Yaskawa INFORM job: STAR.JBI

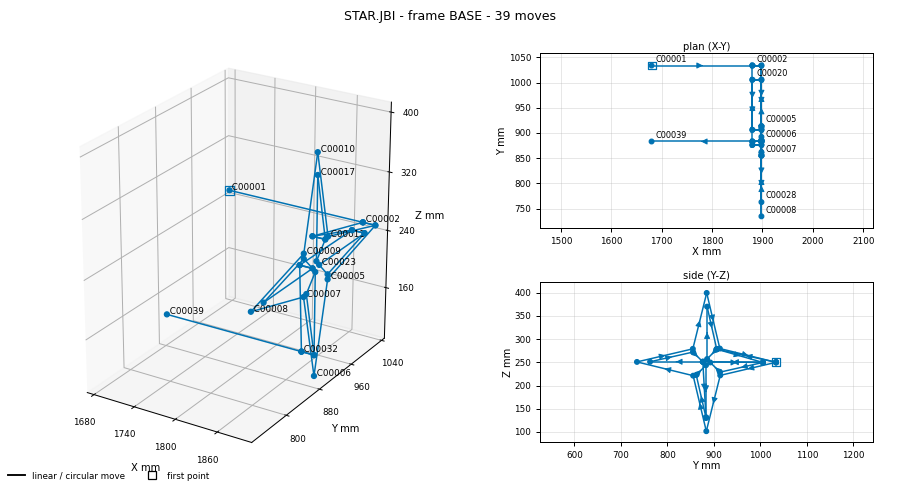
[picture p0: tool path of STAR.JBI in frame BASE, 39 of 40 moves have a stored position in this frame; points joined in program order, loops and branches not executed]
/JOB
//NAME STAR
//POS
///NPOS 40,0,0,0,0,0
///TOOL 9
///POSTYPE PULSE
///PULSE
C00000=38,23,-28,-44,61,-64
///TOOL 9
///POSTYPE BASE
///RECTAN
///RCONF 1,0,0,0,0,0,0,0
C00001=1680.000,1033.806,249.952,-90.00,-0.00,-90.00
C00002=1880.000,1033.806,249.952,-90.00,-0.00,-90.00
C00003=1880.000,1033.806,249.952,-90.00,-0.00,-90.00
C00004=1898.000,1033.806,249.952,-90.00,-0.00,-90.00
C00005=1898.000,913.725,221.863,-90.00,-0.00,-90.00
C00006=1898.000,883.747,101.722,-90.00,-0.00,-90.00
C00007=1898.000,855.472,221.186,-90.00,-0.00,-90.00
C00008=1898.000,734.538,250.798,-90.00,-0.00,-90.00
C00009=1898.000,854.791,278.888,-90.00,-0.00,-90.00
C00010=1898.000,884.598,399.198,-90.00,-0.00,-90.00
C00011=1898.000,912.873,279.564,-90.00,-0.00,-90.00
C00012=1898.000,1033.806,249.952,-90.00,-0.00,-90.00
C00013=1880.000,1033.806,249.952,-90.00,-0.00,-90.00
C00014=1880.000,906.230,278.211,-90.00,-0.00,-90.00
C00015=1898.000,906.230,278.211,-90.00,-0.00,-90.00
C00016=1898.000,885.450,257.059,-90.00,-0.00,-90.00
C00017=1898.000,885.450,369.755,-90.00,-0.00,-90.00
C00018=1898.000,906.230,278.211,-90.00,-0.00,-90.00
C00019=1880.000,906.230,278.211,-90.00,-0.00,-90.00
C00020=1880.000,1005.532,249.614,-90.00,-0.00,-90.00
C00021=1898.000,1005.532,249.614,-90.00,-0.00,-90.00
C00022=1898.000,913.384,228.801,-90.00,-0.00,-90.00
C00023=1898.000,892.263,249.614,-90.00,-0.00,-90.00
C00024=1898.000,1005.532,249.614,-90.00,-0.00,-90.00
C00025=1880.000,1005.532,249.614,-90.00,-0.00,-90.00
C00026=1880.000,876.252,251.137,-90.00,-0.00,-90.00
C00027=1898.000,876.252,251.137,-90.00,-0.00,-90.00
C00028=1898.000,762.813,251.137,-90.00,-0.00,-90.00
C00029=1898.000,854.961,271.950,-90.00,-0.00,-90.00
C00030=1898.000,876.252,251.137,-90.00,-0.00,-90.00
C00031=1880.000,876.252,251.137,-90.00,-0.00,-90.00
C00032=1880.000,883.065,130.996,-90.00,-0.00,-90.00
C00033=1898.000,883.065,130.996,-90.00,-0.00,-90.00
C00034=1898.000,862.115,222.540,-90.00,-0.00,-90.00
C00035=1898.000,883.065,243.691,-90.00,-0.00,-90.00
C00036=1898.000,883.065,130.996,-90.00,-0.00,-90.00
C00037=1880.000,883.065,130.996,-90.00,-0.00,-90.00
C00038=1880.000,883.065,130.996,-90.00,-0.00,-90.00
C00039=1680.000,883.065,130.996,-90.00,-0.00,-90.00
//INST
///DATE 2026/10/26 01:19
///COMM Generated using RoboDK
///ATTR SC,RW,RJ
///GROUP1 RB1
NOP
'Using Tool3 (targets wrt base
'):
'1900.0,883.5,250.0,90.0,0.0,-
'90.0
'Setting Tool 9 (USER - CONE -
' 10MM  X  45 DEG):
SETE P00095 (1) 0
SETE P00095 (2) 0
SETE P00095 (3) 85000
SETE P00095 (4) 0
SETE P00095 (5) 0
SETE P00095 (6) 0
SETTOOL TL#(9) P00095
'hide BALL END - 10MM
'show USER - CONE - 10MM  X  4
'5 DEG
MSG "/ ALPHACAM DRAWING FILE -"
MSG " ROBOTAPT"
MSG "/ NC CODE FILE - ROBOTAPT"
MSG ".apt"
MSG "/ POST-PROCESSED FOR APT-"
MSG "CL DATA"
MSG "/ CREATED - 26 NOV 18"
MSG "/ PROGRAMMED BY ALPHACAM"
MSG "/ USER - CONE - 10MM  X  "
MSG "45 DEG"
MOVJ C00000 VJ=50.00
MOVL C00001 V=1000.0
MOVL C00002 V=1000.0
CALL JOB:SPINDLE
MOVL C00003 V=1000.0
MOVL C00004 V=160.0
MOVL C00005 V=160.0
MOVL C00006 V=160.0
MOVL C00007 V=160.0
MOVL C00008 V=160.0
MOVL C00009 V=160.0
MOVL C00010 V=160.0
MOVL C00011 V=160.0
MOVL C00012 V=160.0
MOVL C00013 V=1000.0
MOVL C00014 V=1000.0
MOVL C00015 V=160.0
MOVL C00016 V=80.0
MOVL C00017 V=160.0
MOVL C00018 V=160.0
MOVL C00019 V=1000.0
MOVL C00020 V=1000.0
MOVL C00021 V=160.0
MOVL C00022 V=80.0
MOVL C00023 V=160.0
MOVL C00024 V=160.0
MOVL C00025 V=1000.0
MOVL C00026 V=1000.0
MOVL C00027 V=160.0
MOVL C00028 V=80.0
MOVL C00029 V=160.0
MOVL C00030 V=160.0
MOVL C00031 V=1000.0
MOVL C00032 V=1000.0
MOVL C00033 V=160.0
MOVL C00034 V=80.0
MOVL C00035 V=160.0
MOVL C00036 V=160.0
MOVL C00037 V=1000.0
CALL JOB:SPINDLE
MOVL C00038 V=1000.0
MOVL C00039 V=1000.0
END
